{attribute 'qualified_only'}
{attribute 'strict'}
{attribute 'to_string'}
TYPE E_PolarIIChamberSwitchModeAfterFinish :
(
	NoChange := 0,
	DryRun := 1,
	Auto := 2
) UINT;
END_TYPE

(* stored: Version 1.1.0.1, ProductVersion 3.1.4026.18
   DUT E_PolarIIChamberSwitchModeAfterFinish: Id {14000000-0000-0000-0000-000000000003} *)
